Staubli VAL3: io.pjx

--- io.pjx ---
parameters version=s6.0 stackSize=0 millimeterUnit=true
data file=io.dtx

--- io.dtx ---

